Universal Robots URScript: T012_codellama_34b-instruct-q4_K_M_baseline_rep1.urscript

urscript

def program():
    # Home the robot
    movej(p[0.0, 0.0, 0.0, 0.0, 0.0, 0.0], a=200.0, v=200.0)

    # Approach spot 1
    movel(p[0.0, 0.0, 0.0, 0.0, 0.0, 0.0], a=200.0, v_tcp=200.0)

    # Descend to spot 1
    movel(p[0.0, 0.0, 0.0, 0.0, 0.0, 0.0], a=80.0, v_tcp=80.0)

    # Lift from spot 1
    movel(p[0.0, 0.0, 0.0, 0.0, 0.0, 0.0], a=150.0, v_tcp=150.0)

    # Move to spot 2
    movel(p[0.0, 0.0, 0.0, 0.0, 0.0, 0.0], a=200.0, v_tcp=200.0)

    # Approach spot 2
    movel(p[0.0, 0.0, 0.0, 0.0, 0.0, 0.0], a=200.0, v_tcp=200.0)

    # Descend to spot 2
    movel(p[0.0, 0.0, 0.0, 0.0, 0.0, 0.0], a=80.0, v_tcp=80.0)

    # Lift from spot 2
    movel(p[0.0, 0.0, 0.0, 0.0, 0.0, 0.0], a=150.0, v_tcp=150.0)

    # Move to spot 3
    movel(p[0.0, 0.0, 0.0, 0.0, 0.0, 0.0], a=200.0, v_tcp=200.0)

    # Approach spot 3
    movel(p[0.0, 0.0, 0.0, 0.0, 0.0, 0.0], a=200.0, v_tcp=200.0)

    # Descend to spot 3
    movel(p[0.0, 0.0, 0.0, 0.0, 0.0, 0.0], a=80.0, v_tcp=80.0)

    # Lift from spot 3
    movel(p[0.0, 0.0, 0.0, 0.0, 0.0, 0.0], a=150.0, v_tcp=150.0)

    # Move to home position
    movej(p[0.0, 0.0, 0.0, 0.0, 0.0, 0.0], a=200.0, v=200.0)

end
